TYPE ST_Prod_Recipe :
STRUCT
	
// General
	Description				: STRING(30);
	prodType				: E_Prod_Type;
	Temperature				: REAL:=4.0;
	
	StirrerDissolving		: ST_Prod_Param_Stirrer;
	StirrerProduction		: ST_Prod_Param_Stirrer;
	StirrerStorage			: ST_Prod_Param_Stirrer;

	ExpirationTime			: TIME:=T#12H;
	Conductivity			: REAL;		// mSimons

	
// Water
	WaterPercentage			: REAL;
	ExpirationTime_Water	: TIME:=T#2D;
	
// Line	
	ExpirationTime_Line			: TIME:=T#24H;
	ExpirationTime_Line_Stby	: TIME:=T#2H;
	
// Component
	arr_Component			: ARRAY [1..g_Prod.cMaxCompInProduct] OF ST_Prod_Ingredient;
	
// Water push to triblender color(Blood)
	Weight_to_Collect		: REAL:=60; // Kg
	Weight_to_Drain			: REAL:=200; // Kg
	Conductivity_limit		: REAL; //mSimons
	
	
	FlowRate_Production		: REAL:=800; //RPM
	FlowRate_WaterPushing	: REAL:=800; //RPM
	FlowRate_Storage		: REAL:=800; //RPM
	
	eFilling_Mode			: E_Filling_Mode;
	BinWeight				: REAL:=200.0;	//kg
	BinWeightTolerance		: REAL:=0.5;	//kg




END_STRUCT
END_TYPE

(* stored: Version 1.1.0.1, ProductVersion 3.1.4024.15
   DUT ST_Prod_Recipe: Id {30f796b6-4ad6-4488-9821-178c2ff4e475} *)
